(* IEC 61131-3 sources: CodesysTools/tests/samples, 14 files *)

(* ---- naming_noprefix.st ---- *)
//{attribute 'noprefix'}
{attribute 'pack_mode' := '1'}
TYPE tMbUnion :
UNION
    b  : tMbState;  //For Bit Access
    dw : DWord;     //For DoubleWord Access
    w2 : WORD;
    Raw : INT;
    foo : INT;
END_UNION
END_TYPE

(* ---- naming_union.st ---- *)
{attribute 'pack_mode' := '1'}
TYPE tMbUnion :
UNION
    b  : tMbState;  //For Bit Access
    dw : DWord;     //For DoubleWord Access
    w2 : WORD;
    Raw : INT;
    foo : INT;
END_UNION
END_TYPE

(* ---- decl_init.st ---- *)
FUNCTION_BLOCK FB_X
VAR
    sValve:tValve(bOpen:=TRUE, iMax:=10, rGain := 1.5);   // valve
    sb : BOOL;
    sName : STRING(80) := 'x';
    {attribute 'a'} sOther : tOther := (iA:=1,iB:=2);
    saArr : ARRAY[1..2] OF INT := [1,2];
END_VAR
sb := TRUE;

(* ---- general.st ---- *)
FUNCTION_BLOCK fb_Motor EXTENDS fb_Base
VAR_INPUT
bStart:BOOL;   // start command
  bStop : BOOL:=FALSE; (* stop *)
nSpeedSetpoint:INT;
END_VAR
var
tonDelay:TON;
aBuffer : ARRAY [1..10] OF REAL;
sName:STRING(80):='Motor $'A$'';
iState : INT;
dtStart:DT:=DT#2024-01-01-12:30:00;
pIn AT %IX0.1:BOOL;
end_var

(* main logic *)
if bStart and not bStop then
iState:=1;
elsif bStop then
iState := 0;
else
   x:=-5+y*(3-z);
end_if

case iState of
0:
tonDelay(IN:=FALSE,PT:=T#2S);
1,2:   tonDelay(IN:=TRUE,
PT:=T#5s);
IF tonDelay.Q THEN
iState:=E_State#Running;
END_IF
-1: ;
else
iState:=0;
end_case

FOR i:=1 TO 10 BY 1 DO
aBuffer[i]:=INT_TO_REAL(i)*1.5E3;
END_FOR
REPEAT
i:=i+1;
UNTIL i>5
END_REPEAT;
END_FUNCTION_BLOCK

TYPE ST_Data :
STRUCT
a:INT; // first
longName : LREAL := 1.0;
END_STRUCT
END_TYPE

PROGRAM Main
VAR
    i:INT; (* loop counter *)
    rTemperatureActual : REAL := 20.5; // measured
    bAlarm:BOOL;
END_VAR
i:=0; // reset
rTemperatureActual:=rTemperatureActual+0.1;
bAlarm := rTemperatureActual>80.0;   // high temp
THIS^.x:=1;
END_PROGRAM

(* ---- naming.st ---- *)
VAR_GLOBAL
    gbAlarm : BOOL;
    bAlarm2 : BOOL;
    iStart AT %IX0.0 : BOOL;
    ibStop AT %IX0.1 : BOOL;
    qbLamp AT %QX0.0 : BOOL;
END_VAR
VAR_GLOBAL CONSTANT
    gciMax : INT := 10;
    MAX_N : INT := 5;
END_VAR
FUNCTION_BLOCK fbMotor
VAR_INPUT
    ibReset : BOOL;
    nSpeed : INT;
    ixEnable, bRun : BOOL;
    iAxis : ST_Axis;
END_VAR
VAR_OUTPUT
    qrSpeed : REAL;
    qlrPos : LREAL;
END_VAR
VAR_IN_OUT
    iqData : ST_Data;
END_VAR
VAR
    sbReset : BOOL;
    tonDelay : TON;
    sTimer : TON;
    aBuf : ARRAY[1..10] OF REAL;
    srBuf2 : ARRAY[1..10] OF REAL;
    sudiCount : UDINT := 0;
    sString : STRING(80);
    ssName : STRING(80);
    sdtStamp : DT;
END_VAR
VAR CONSTANT
    ciLimit : INT := 3;
END_VAR
VAR_TEMP
    ttElapsed : TIME;
    tData : ST_Data;
END_VAR
END_FUNCTION_BLOCK
FUNCTION fcAdd : INT
VAR
    tiX : INT;
    siY : INT;
END_VAR
END_FUNCTION
TYPE ST_Data :
STRUCT
    bOk : BOOL;
    rVal : REAL;
    value : INT;
    Sub : ST_Sub;
END_STRUCT
END_TYPE

(* ---- naming_block_skip.st ---- *)
TYPE tA :
STRUCT //{attribute 'noprefix'}
    Alpha : INT;
    Beta : BOOL;
END_STRUCT
END_TYPE
TYPE tB :
STRUCT
    Gamma : INT;
END_STRUCT
END_TYPE
FUNCTION_BLOCK FB_X
VAR (* {attribute 'noprefix'} *)
    Free : INT;
END_VAR
VAR
    Checked : INT;
END_VAR
END_FUNCTION_BLOCK

(* ---- naming_prefixes.st ---- *)
FUNCTION_BLOCK FB_T
VAR
    kMaxSize : INT := 3;
    vSpeed : REAL;
    mValue : BOOL;
    mode : INT;
    kmax : INT;
    m : INT;
    sbOk : BOOL;
    sb2Valve : BOOL;
    sbValve2 : BOOL;
    k2Max : INT;
    sb_x : BOOL;
    k : INT;
    k_1 : INT;
    v : INT;
    smRot : REAL;
    tmRot : REAL;
    svPos : REAL;
    tvPos2 : REAL;
    tmp : REAL;
    gmRot : REAL;
END_VAR
END_FUNCTION_BLOCK

(* ---- naming_types.st ---- *)
FUNCTION_BLOCK FB_T
VAR
    Start : TOD;
    Data : ST_Data;
    aData : ARRAY[0..3] OF ST_Data;
    Other : ST_Other;
    Flag : BOOL;
END_VAR
END_FUNCTION_BLOCK

(* ---- region_attributes.st ---- *)
FUNCTION_BLOCK fb_Motor
VAR_INPUT
    bStart:BOOL;   // start command
        {attribute 'hide'}
    bInternalFlagLongName : BOOL:=FALSE; (* stop *)
  {attribute 'hide'}   nCnt:LINT;
END_VAR
var_output
x:lreal; // out
end_var
REGION Motor If control
if bStart then
iState:=1; // run
elsif bStop then
iCounterValue:=0;
else
   x:=-5;
end_if
END_REGION
for i:=1 to 10 do
aBuffer[i]:=i; // fill
end_for
END_FUNCTION_BLOCK

(* ---- spelling.st ---- *)
// This valve is wrong, the wrod is spelled wrong
(* Valves and unhappy workers check the lines *)
FUNCTION_BLOCK FB_Valve
VAR
    sbOpen : BOOL;  // The valve colour: a PLC flag with a mispelling
    sbValveOk : BOOL;  // valvs of London and tMbState and sValve
END_VAR
// sbOpen := TRUE;  commented out code is skipped
// See https://example.com/wrodd and file.txt for details
sbOpen := TRUE; // Worke it, e.g. unworkers and valveed
(* Multi
   line commment
   second: chek the line *)
// {attribute 'noprefix'}
// arbeidsbord og ventilbord, løs og ære, feilstavet ventilbrod
END_FUNCTION_BLOCK

(* ---- terminal_codes.st ---- *)
FUNCTION_BLOCK FB_Valve
VAR_INPUT
    R : BOOL;
    BA1 : BOOL;
    XE : BOOL;
    START_CMD : BOOL;
    BZ : BOOL;
    QA : BOOL;
    Start : BOOL;
    ibReset : BOOL;
END_VAR
VAR_OUTPUT
    YH : BOOL;
    qbOpen : BOOL;
END_VAR
VAR
    START : BOOL;
END_VAR
END_FUNCTION_BLOCK

(* ---- calls.st ---- *)
PROGRAM Main
VAR
    sTimer : TON;
    sbStart : BOOL;
    sbDone : BOOL;
    stElapsed : TIME;
    srX : REAL;
END_VAR
sbStart:=TRUE;
sTimer(IN:=sbStart, PT:=T#5S, // time
       Q=>sbDone, ET=>stElapsed);   // done
IF sbStart THEN
  aFb[1].Run(Execute := TRUE);
  srX := LIMIT(0.0, srX, 10.0);
  F_Calc(srX);
END_IF
srX := a +
  F(b := 1);
sTimer(
// comment line
IN:=sbStart);
END_PROGRAM

(* ---- functions.st ---- *)
PROGRAM P
VAR
    sR : LREAL;
END_VAR
sR := ABS(x) + sin (y) + INT_TO_REAL(i) + to_int(r) + MAX(a, b) + st.Len + LIMIT(0, a, 5);
sR := stX.max;
sR := ltime_to_lreal(a) + to_dword(c) + TRUNC_INT(d) + TOD_TO_TIME(f);

(* ---- typed_literals.st ---- *)
PROGRAM P
VAR
    sT : LTIME := ltime#1s;
    sB : INT := INT#5;
END_VAR
sT := tod#12:00:00; sB := 16#FF; sT := T#5s; sT := dint#3;
